(* IEC 61131-3 sources: plcassist-cli/packages/volt-lsp-iec/test-corpus/lenze-mid/Device/Plc Logic/Application/A70_MachineModuleSources/MM_MachineControl/02_subMain, 11 files *)

(* ---- SidecorrectionCalculation.fun ---- *)
FUNCTION SidecorrectionCalculation
VAR_INPUT
	iAnalogInputValue						: INT;
	iSetpoint								: INT;
	iCorrectionScale						: REAL;
	iLightValue								: INT;
	iDarkValue								: INT;
	iNoWrapperOffsetPercentage01Perc		: INT; //test5

END_VAR
VAR_OUTPUT
	oIntPercentage							: INT;
	oRealPercentage							: REAL;
	oCorrectionValue						: REAL;
	oDeviationNoWrapper						: REAL;
END_VAR
VAR

	tRealMeasuredValue						: REAL;
	tRealPercentage							: REAL;
	tRealSetpoint							: REAL;
	tWhiteValue								: DINT;
	tBrownValue								: DINT;
	tWidthLight_Dark						: DINT;
	tRealWidthLight_Dark					: REAL;
	tMeasuredWithOffset						: REAL;
	tRealBrownValue							: REAL;
	tRealNoWrapperOffsetPercentage			: REAL;

END_VAR

//Read out values for light and dark
tWhiteValue:=MOVE(iLightValue);
tBrownValue:=MOVE(iDarkValue);

//Calculate difference between light and dark value (light will be higher than dark)
tRealWidthLight_Dark:=TO_REAL(tWhiteValue-tBrownValue);
tRealBrownValue:=TO_REAL(tBrownValue);

//Measured value compensated with offset
tRealMeasuredValue:=TO_REAL(iAnalogInputValue);
tMeasuredWithOffset:=tRealMeasuredValue-tRealBrownValue;

//Calculation of the percentage
//"Measured value"/ Bandwidth
IF tRealWidthLight_Dark=0 THEN
	tRealWidthLight_Dark:=10;

END_IF
oRealPercentage:=(tMeasuredWithOffset/tRealWidthLight_Dark)*100;
oIntPercentage:=TO_INT(oRealPercentage);

//Calculation of the fault
//(act - set) * "correction scale"
tRealSetpoint:=TO_REAL(iSetpoint);
oCorrectionValue:=(oRealPercentage-tRealSetpoint)*iCorrectionScale;

//No wrapper detection
tRealNoWrapperOffsetPercentage:=TO_REAL(iNoWrapperOffsetPercentage01Perc);
oDeviationNoWrapper:=TO_INT(tRealNoWrapperOffsetPercentage*(tRealWidthLight_Dark/1000));

END_FUNCTION

(* ---- SpeedCalculationTrayfiller.fun ---- *)
FUNCTION SpeedCalculationTrayfiller
VAR_INPUT
END_VAR
VAR
	tInt: INT;
	tBool: BOOL;
END_VAR

NETWORK 0 LD TITLE: "NETWORK 1: Write setpoint speed in DB"
  // The speed of the trayfiller has to be higher then the speed of the dryer. In this way there is always an empty space at the startpostition of the trayfiller.
  LET en1 := ;
  IF en1 THEN tInt := (Mach1_Data.Drives.FeedForwardADS.Control.AutoSpeed + 30); END_IF
  LET en2 := en1;
  IF en2 THEN Mach1_Data.Drives.FeedForwardATF.Control.AutoSpeed := MOVE(tInt); END_IF
END_NETWORK
NETWORK 1 LD TITLE: "NETWORK 2: Activation + Runtime guard feed forward dryer/trayfiller"
  // Runtime calculation:
  // 1 cycle = 60s/rpm
  // speed = in 0.1 rpm -> 60s = 600 1/10s
  //
  // -> 1 cycle = 600/speed01
  // DINT cannot calculate this 600/1000 = 0.1 -> DINT=0
  // First multiply by 1000 (s -> ms)
  // 1cycle = (600*1000)/speed1
  // To give a little margin: add 500ms
  LET en1 := (Mach1.Genflags.DelayAfterSTO AND Mach1_Data.Drives.FeedForwardATF.Control.StartAuto AND NOT LST_InputsOutputs.I133_3_PROX_zero_position_transport_ATF);
  IF en1 THEN (Mach1_Data.Drives.FeedForwardATF.Control.AutoSpeed >= 10); END_IF
  Mach1.GenFlags.StopDriveDirect S= RuntimeGuard_V5_1_100(Mach1_Alarms, (Mach1_AuxData.TrayfillerActive AND Mach1_MIDS.IDB_TrayFiller.oFeedForwardMotor AND Mach1.Genflags.DelayAfterSTO AND (Mach1_AuxData.AllDrivesHomed OR NOT Mach1_AuxData.TrayfillerActive)), LST_General.AlwaysOff, en1, T#10S, Mach1.GenFlags.StartFlag, Mach1_Alarms.Alm051, Mach1.GenFlags.MinorAlarm, Mach1_AuxData.IEC_TIMERS.RuntimeGuardFeedforwardTrayfiller, oForwardGuarded => Mach1_Data.Drives.FeedForwardATF.Control.StartAuto);
END_NETWORK

END_FUNCTION

(* ---- Servo_LimitJog.fb ---- *)
FUNCTION_BLOCK Servo_LimitJog
VAR_INPUT
	iServoStatus 	: sUDT_ServoComm_Drive_Status;
	iServoControl 		: sUDT_ServoComm_Drive_Control;
END_VAR
VAR_OUTPUT
	oServoControl 		: sUDT_ServoComm_Drive_Control;
END_VAR
VAR
END_VAR
VAR_IN_OUT
	ioUDT_ServoDrive			: UDT_ServoDrive;
	ioUDT_JogLimitFree			: UDT_ServoJogLimitFree;
END_VAR

NETWORK 0 LD TITLE: "NETWORK 3 (p1): Check for limit switch"
  ioUDT_JogLimitFree.Status.Limit_Left_OK := iServoStatus.Spare1;
END_NETWORK
NETWORK 1 LD TITLE: "NETWORK 3 (p2): Check for limit switch"
  ioUDT_JogLimitFree.Status.Limit_Right_OK := iServoStatus.Spare2;
END_NETWORK
NETWORK 2 LD TITLE: "COPY previous control word to current controlword"
  LET en1 := ;
  IF en1 THEN
  EXECUTE
oServoControl:=iServoControl;
  END_EXECUTE
  END_IF
END_NETWORK
NETWORK 3 LD TITLE: "NETWORK 4 (p1): ControlToFreeLimitSwitches"
  oServoControl.Spare1 := (ioUDT_JogLimitFree.Status.Limit_Left_OK AND ioUDT_JogLimitFree.Control.Jog_LimitToLeft);
END_NETWORK
NETWORK 4 LD TITLE: "NETWORK 4 (p2): ControlToFreeLimitSwitches"
  oServoControl.Spare2 := (ioUDT_JogLimitFree.Status.Limit_Right_OK AND ioUDT_JogLimitFree.Control.Jog_LimitToRight);
END_NETWORK

END_FUNCTION_BLOCK

(* ---- WSM.fb ---- *)
FUNCTION_BLOCK WSM
VAR_INPUT
	EN: BOOL;
	iGenflags : UDT_GeneralFlags;
	iInit: BOOL;
	iTest_Prod: BOOL;
	iCleaning: BOOL;
	iBunchPresent: BOOL;
	iWrapperPresentForLeafCarrier: BOOL;
	iPhotocellWrapper: BOOL;
	iWaterLevelSensor: BOOL;
	iTakeOverCycle: BOOL;
	iTimeOutSupplyWrapper: TIME;
	iSprayTime: TIME;
	iDelayContSpraying: TIME;
	iScreenForOperatorSettingsActivated: BOOL;
	iManualSprayCycleReset: BOOL;
	iManualSprayCycleStart: BOOL;
	iManualSprayCycleStop: BOOL;
	iMaxNumberOfSprayPulses: INT;

END_VAR
VAR_OUTPUT
	ENO: BOOL;
	oVentilationMotor: BOOL;
	oPositionMotor: BOOL;
	oWindingMotor: BOOL;
	oSprayingValve: BOOL;
	oWaterLevelValve: BOOL;
	oFaultWaitingForWrapper: BOOL;
	oFaultNoWrapper: BOOL;
	oFaultPhotocellWrapper : BOOL;
END_VAR
VAR
	stOSN_TakeOverCycle: F_TRIG;
	TMR_TimeOutSupply: TON;
	TMR_TimeOutPhotocell: TON;
	stRePositionMotor: R_TRIG;
	stSprayCycleActive: BOOL;
	TMR_DelayContinuousSpraying: TON;
	TMR_SprayTime: TON;
	stManualSprayCycleStarted: BOOL;

	TMR_ManualSprayCycleIdle: TON;

END_VAR

VAR_IN_OUT
	ioEnableSpraying: BOOL;
	ioManualSprayCycleActualCount: INT;
	ioManualStartSupply: BOOL;
END_VAR
VAR RETAIN PERSISTENT
	stRestposition: BOOL;
	stSupplyWrapper: BOOL;
	stWrapperPresent: BOOL;
	stNoWrapper: BOOL;
	stPhotocellWrapperFault: BOOL;
	stFeedForward: BOOL;
END_VAR

NETWORK 0 LD TITLE: "DONE Network 2: State: Initialise"
  LET g8 := (iInit OR NOT iTest_Prod OR iCleaning OR ioManualStartSupply);
  stRestposition S= g8;
  LET g1 := g8;
  stSupplyWrapper R= g1;
  stWrapperPresent R= g1;
  stNoWrapper R= g1;
  stPhotocellWrapperFault R= g1;
END_NETWORK
NETWORK 1 LD TITLE: "DONE Network 3: State: Restposition"
  LET g1 := (stOSN_TakeOverCycle(CLK := iTakeOverCycle) AND stWrapperPresent);
  stRestposition S= g1;
  stWrapperPresent R= g1;
END_NETWORK
NETWORK 2 LD TITLE: "DONE Network 4: State: Supply wrapper"
  LET g1 := ((stRestposition AND ((iTest_Prod AND NOT iCleaning AND iBunchPresent AND NOT iTakeOverCycle AND (iGenFlags.RunMan OR iGenFlags.RunAuto)) OR ioManualStartSupply)) OR (stNoWrapper AND iGenFlags.StartFlag) OR (stPhotocellWrapperFault AND iGenFlags.StartFlag));
  stSupplyWrapper S= g1;
  stRestposition R= g1;
  stNoWrapper R= g1;
  stPhotocellWrapperFault R= g1;
  ioManualStartSupply R= g1;
END_NETWORK
NETWORK 3 LD TITLE: "DONE Network 5: State: Wrapper Present"
  LET g15 := (iWrapperPresentForLeafCarrier AND stSupplyWrapper);
  stWrapperPresent S= g15;
  LET en1 := g15;
  IF en1 THEN HMI_Var.Mach1.PRDWrapCurrentCntr := (1 + HMI_Var.Mach1.PRDWrapCurrentCntr); END_IF
  LET en2 := g15;
  IF en2 THEN HMI_Var.Mach1.PRDWrapDayCounter := (1 + HMI_Var.Mach1.PRDWrapDayCounter); END_IF
  stSupplyWrapper R= g15;
END_NETWORK
NETWORK 4 LD TITLE: "DONE Network 6: State: No Wrapper"
  LET g1 := TMR_TimeOutSupply(IN := (stSupplyWrapper AND stFeedForward), PT := iTimeOutSupplyWrapper);
  stNoWrapper S= g1;
  stSupplyWrapper R= g1;
END_NETWORK
NETWORK 5 LD TITLE: "DONE Network 7: State: Photocell wrapper fault"
  LET g1 := TMR_TimeOutPhotocell(IN := (stSupplyWrapper AND stFeedForward AND iPhotocellWrapper), PT := T#10S);
  stPhotocellWrapperFault S= g1;
  stSupplyWrapper R= g1;
END_NETWORK
NETWORK 6 LD TITLE: "DONE Network 8: Faults"
  LET g21 := True;
  oFaultWaitingForWrapper := (g21 AND stSupplyWrapper AND iTakeOverCycle);
  oFaultNoWrapper := (g21 AND stNoWrapper);
  oFaultPhotocellWrapper := (g21 AND stPhotocellWrapperFault);
END_NETWORK
NETWORK 7 LD TITLE: "DONE Network 9: Ventilation motor"
  oVentilationMotor := (iGenFlags.EnableAuxDrive AND iTest_Prod AND NOT iCleaning);
END_NETWORK
NETWORK 8 LD TITLE: "DONE Network 10:"
  LET g23 := (iGenFlags.EnableAuxDrive AND stSupplyWrapper AND NOT iGenFlags.StopFlag);
  stFeedForward := g23;
  oPositionMotor := g23;
END_NETWORK
NETWORK 9 LD TITLE: "DONE Network 11: Winding motor"
  oWindingMotor := (iGenFlags.EnableAuxDrive AND NOT iGenFlags.StopFlag AND iTest_Prod AND NOT iCleaning);
END_NETWORK
NETWORK 10 LD TITLE: "DONE Network 12: Start spray cycle"
  LET g46 := stFeedForward;
  stSprayCycleActive S= stRePositionMotor(CLK := g46);
  stSprayCycleActive S= TMR_DelayContinuousSpraying(IN := g46, PT := iDelayContSpraying);
END_NETWORK
NETWORK 11 LD TITLE: "DONE Network 13: Timing spray cycle"
  stSprayCycleActive R= (TMR_SprayTime(IN := stSprayCycleActive, PT := iSprayTime) AND NOT TMR_DelayContinuousSpraying.Q);
END_NETWORK
NETWORK 12 LD TITLE: "DONE Network 14: Spraying valve"
  oSprayingValve := (ioEnableSpraying AND stSprayCycleActive);
END_NETWORK
NETWORK 13 LD TITLE: "DONE Network 15: Automatic trigger of water"
  ioEnableSpraying S= (FALSE AND iGenFlags.EnablePneumEStop AND iWrapperPresentForLeafCarrier AND iTest_Prod AND NOT iCleaning);
END_NETWORK
NETWORK 14 LD TITLE: "DONE Network 16: Water level control"
  oWaterLevelValve := (ioEnableSpraying AND iWaterLevelSensor);
END_NETWORK
NETWORK 15 LD TITLE: "DONE Network 17: Manual spray cycle"
  LET g45 := iScreenForOperatorSettingsActivated;
  LET en1 := (g45 AND iManualSprayCycleReset);
  IF en1 THEN ioManualSprayCycleActualCount := MOVE(0); END_IF
  LET en2 := (g45 AND iGenFlags.EnablePneumEStop AND (iManualSprayCycleStart OR stManualSprayCycleStarted) AND NOT iManualSprayCycleStop AND NOT iManualSprayCycleReset);
  IF en2 THEN stManualSprayCycleStarted := (ioManualSprayCycleActualCount < iMaxNumberOfSprayPulses); END_IF
  LET en3 := TMR_ManualSprayCycleIdle(IN := (g45 AND stManualSprayCycleStarted AND NOT stSprayCycleActive), PT := T#300MS);
  IF en3 THEN ioManualSprayCycleActualCount := (ioManualSprayCycleActualCount + 1); END_IF
  stSprayCycleActive S= en3;
END_NETWORK
NETWORK 16 LD TITLE: "DONE Network 18: SAVE RLO"
  ENO := EN;
END_NETWORK

END_FUNCTION_BLOCK

(* ---- AHWF.prg ---- *)
PROGRAM AHWF
VAR
	tFaultWaitingForWrapper : BOOL;
	tFaultNoWrapper: BOOL;
	tFaultPhotocellWrapper: BOOL;
	tStartFastWinding: BOOL;
	tSupplyWrapper: BOOL;
	tSprayingValve: BOOL;
	ttest: BOOL;
	R_TrigStartPos: R_TRIG;
END_VAR

VAR
	IDB_WSM: WSM;
END_VAR

NETWORK 0 LD TITLE: "Network 1: Detection of wrapper (set and reset)"
  LET g10 := True;
  Mach1_AuxData.MemWrapperPassedUnderTheSensor S= (g10 AND LST_InputsOutputs.I101_0_Wrapper_present);
  LET g1 := (g10 AND NOT LST_InputsOutputs.I101_0_Wrapper_present AND Mach1_AuxData.MemWrapperPassedUnderTheSensor);
  Mach1_AuxData.MemWrapperPresentForLeafCarrier S= g1;
  Mach1_AuxData.MemWrapperDetected_ResetLimitedSpeed S= g1;
  LET en1 := g10;
  IF en1 THEN Mach1_AuxData.CamControls.TakeOverCycleStopPulse_CP.Start := MOVE(Mach1_Data.CamControls.TakeOverCycle_C.Stop); END_IF
  LET g2 := fc_CamC_CP_UDT(en1, HMI_Var.Mach1.Position, Mach1.GenFlags.Rotflag, Mach1_AuxData.CamControls.TakeOverCycleStopPulse_CP);
  Mach1_AuxData.MemWrapperPresentForLeafCarrier R= g2;
  Mach1_AuxData.MemWrapperPassedUnderTheSensor R= g2;
END_NETWORK
NETWORK 1 LD
  LET g1 := R_TrigStartPos(CLK := HMI_Var.HMI_AHWF_StartPos);
  Mach1_AuxData.MemWrapperPresentForLeafCarrier R= g1;
  Mach1_AuxData.MemWrapperPassedUnderTheSensor R= g1;
END_NETWORK
NETWORK 2 LD TITLE: "Network 2: FB for DTA"
  LET i1 := fc_dinttotime(Mach1_Data.Timers.TimeOutSupplyWrapper,2);
  LET i2 := fc_dinttotime(Mach1_Data.Timers.SprayPulseWidth,2);
  LET i3 := fc_dinttotime(Mach1_Data.Timers.DelayContSpraying,2);
  LET en1 := ;
  IF en1 THEN IDB_WSM(iGenflags := Mach1.GenFlags, iInit := LST_General.FirstCycle, iTest_Prod := HMI_Var.Test_Prod, iCleaning := HMI_Var.Btn_Cleaning, iBunchPresent := Mach1_AuxData.ShiftRegister.SR_bunch_present_position_1_JL, iWrapperPresentForLeafCarrier := (Mach1_AuxData.MemWrapperPresentForLeafCarrier AND NOT HMI_Var.HMI_AHWF_fast_winding), iPhotocellWrapper := (LST_InputsOutputs.I101_0_Wrapper_present AND NOT HMI_Var.HMI_AHWF_fast_winding), iWaterLevelSensor := LST_InputsOutputs.I101_3_Water_level_control, iTakeOverCycle := fc_CamC_CC_UDT(True, HMI_Var.Mach1.Position, Mach1_Data.CamControls.TakeOverCycle_C), iTimeOutSupplyWrapper := i1, iSprayTime := i2, iDelayContSpraying := i3, iScreenForOperatorSettingsActivated := Mach1_AuxData.ScreenForOperatorSettingsActivated, iManualSprayCycleReset := HMI_Var.Mach1.SprayReset, iManualSprayCycleStart := HMI_Var.Mach1.SprayStart, iManualSprayCycleStop := HMI_Var.Mach1.SprayStop, iMaxNumberOfSprayPulses := Mach1_Data.Settings.Ints.MaxNumberOfSprayPulses, ioEnableSpraying := HMI_Var.Btn_Spraying, ioManualSprayCycleActualCount := Mach1_Data.Settings.Ints.ActualNumberOfSprayPulses, ioManualStartSupply := HMI_Var.HMI_AHWF_StartPos, oPositionMotor => tSupplyWrapper, oSprayingValve => tSprayingValve, oWaterLevelValve => LST_InputsOutputs.Q101_1_PNV_Waterlevel_control, oFaultWaitingForWrapper => tFaultWaitingForWrapper, oFaultNoWrapper => tFaultNoWrapper, oFaultPhotocellWrapper => tFaultPhotocellWrapper); END_IF
  PneumValveTerminalSMC.Pos1B := (en1 AND Mach1.GenFlags.EnablePneumPressurised AND Mach1_Safety.Status.AllDoorsActuallyClosed AND tSprayingValve AND NOT Mach1_Alarms.Alm011);
END_NETWORK
NETWORK 3 LD TITLE: "Network 3: Wrapper faults"
  Mach1.GenFlags.StopDriveDirect S= (Alarms_V5_1_100(Mach1_Alarms, (Mach1.GenFlags.DelayAfterEmergStop AND HMI_Var.Test_Prod AND NOT HMI_Var.Btn_Cleaning AND tFaultWaitingForWrapper AND Mach1_AuxData.AllDrivesHomed), True, Mach1_Alarms.Alm076, Mach1.GenFlags.Warning) OR Alarms_V5_1_100(Mach1_Alarms, (Mach1.GenFlags.DelayAfterEmergStop AND HMI_Var.Test_Prod AND NOT HMI_Var.Btn_Cleaning AND tFaultNoWrapper AND Mach1_AuxData.AllDrivesHomed), Mach1.GenFlags.StartFlag, Mach1_Alarms.Alm043, Mach1.GenFlags.MinorAlarm) OR Alarms_V5_1_100(Mach1_Alarms, (Mach1.GenFlags.DelayAfterEmergStop AND HMI_Var.Test_Prod AND NOT HMI_Var.Btn_Cleaning AND NOT Mach1_Alarms.Alm045 AND tFaultPhotocellWrapper AND Mach1_AuxData.AllDrivesHomed), Mach1.GenFlags.StartFlag, Mach1_Alarms.Alm045, Mach1.GenFlags.MinorAlarm));
END_NETWORK
NETWORK 4 LD
END_NETWORK
NETWORK 5 LD TITLE: "TODO Network 4:"
  LET g328 := True;
  LET g329 := (g328 AND True);
  LET en1 := (g329 AND TRUE);
  IF en1 THEN Data_Exchange_Motion.FeedForwardWrapper.Control.VelUnit := MOVE(175); END_IF
  LET en2 := en1;
  IF en2 THEN Data_Exchange_Motion.FeedForwardWrapper.Control.DecUnit := MOVE(2000); END_IF
  LET en3 := en2;
  IF en3 THEN Data_Exchange_Motion.FeedForwardWrapper.Control.AccUnit := MOVE(750); END_IF
  LET en4 := en3;
  IF en4 THEN Data_Exchange_Motion.FeedForwardWrapper.Control.TorqueLimit := MOVE(100); END_IF
  LET g330 := (g329 AND HMI_Var.HMI_AHWF_fast_winding);
  tStartFastWinding := Mach1_AuxData.IEC_TIMERS.TON_StartFastWinding(IN := g330, PT := T#200MS);
  LET en5 := g330;
  IF en5 THEN Data_Exchange_Motion.FeedForwardWrapper.Control.VelUnit := MOVE(500); END_IF
  LET i1 := DINT_TO_LREAL(Mach1_Data.Settings.Dints.WrapperStopPosition)/10;
  LET en6 := g328;
  IF en6 THEN Data_Exchange_Motion.FeedForwardWrapper.Control.PosUnit := MOVE(i1); END_IF
  Data_Exchange_Motion.FeedForwardWrapper.Control.StartTouchprobePos := (g328 AND NOT HMI_Var.HMI_AHWF_positioningType AND NOT Mach1_Alarms.Alm056 AND mach1.Genflags.EnableAuxDrive AND (tSupplyWrapper OR tStartFastWinding OR (Data_Exchange_Motion.FeedForwardWrapper.Control.StartTouchprobePos AND NOT Data_Exchange_Motion.FeedForwardWrapper.Status.InPosition)));
  HMI_Var.HMI_AHWF_fast_winding R= Mach1_AuxData.Edge.OSP_StopFlag(CLK := (g328 AND (NOT Mach1_MIDS.FB_Mach1.iStop1 OR NOT Mach1_MIDS.FB_Mach1.iStop2 OR NOT Mach1_MIDS.FB_Mach1.iStop3 OR NOT Mach1_Safety.Status.AllDoorsActuallyClosed OR LST_InputsOutputs.I101_0_Wrapper_present)));
END_NETWORK
NETWORK 6 LD TITLE: "Network 5: Side correction"
  LET en1 := ;
  IF en1 THEN ??? := SideCorrection(); END_IF
END_NETWORK
NETWORK 7 LD TITLE: "Network 6: DTA-alarm: side limit reached"
  Mach1.GenFlags.StopDriveDirect S= (Alarms_V5_1_100(Mach1_Alarms, (Mach1_AuxData.Edge.OSP_LimitDTA_Reached(CLK := (Mach1_AuxData.MIDS_Active AND Mach1.GenFlags.DelayAfterEmergStop AND (NOT Mach1_Data.Drives.SideCorrection_FreeLimit.Status.Limit_Left_OK OR NOT Mach1_Data.Drives.SideCorrection_FreeLimit.Status.Limit_Right_OK))) AND Mach1_AuxData.AllDrivesHomed), Mach1.GenFlags.StartFlag, Mach1_Alarms.Alm057, Mach1.GenFlags.MinorAlarm) OR (LST_General.AlwaysOff AND Alarms_V5_1_100(Mach1_Alarms, (Mach1_AuxData.MIDS_Active AND Mach1.GenFlags.DelayAfterEmergStop AND (NOT Mach1_Data.Drives.SideCorrection_FreeLimit.Status.Limit_Left_OK OR NOT Mach1_Data.Drives.SideCorrection_FreeLimit.Status.Limit_Right_OK) AND Mach1_AuxData.AllDrivesHomed), Mach1.GenFlags.StartFlag, Mach1_Alarms.Alm074, Mach1.GenFlags.Warning)));
END_NETWORK
NETWORK 8 LD TITLE: "Network 7: Alarm: Water receptacle full"
  Mach1.GenFlags.StopDriveDirect S= Alarms_V5_1_100(Mach1_Alarms, (Mach1_AuxData.IEC_TIMERS.WaterReceptacleFull(IN := (Mach1_AuxData.MIDS_Active AND LST_InputsOutputs.I101_3_Water_level_control AND NOT Mach1_Alarms.Alm055), PT := T#5M) AND HMI_Var.Test_Prod AND HMI_Var.Btn_Spraying AND Mach1_AuxData.AllDrivesHomed), Mach1.GenFlags.StartFlag, Mach1_Alarms.Alm055, Mach1.GenFlags.MinorAlarm);
END_NETWORK

END_PROGRAM

(* ---- fc_CheckRegister.prg ---- *)
PROGRAM fc_CheckRegister
VAR
END_VAR

NETWORK 0 LD TITLE: "NETWORK 1: Shift CheckRegister"
  fc_ShiftRegister(db_CheckRegister.Positie);
END_NETWORK
NETWORK 1 LD TITLE: "NETWORK 2: Check for error in dryer"
  fc_CheckNumberOfErrorsRegister(db_CheckRegister.Positie, CTE.posCigarPresentOutfeed, Mach1_Data.Counters.MaxRepetitionNoCigarsDryer.SetValue, oError => db_CheckRegister.CheckRegisterError);
END_NETWORK

END_PROGRAM

(* ---- fc_Visualisation_HMI.prg ---- *)
PROGRAM fc_Visualisation_HMI
VAR_INPUT
END_VAR
VAR
	tbool: BOOL;
END_VAR

NETWORK 0 LD TITLE: "NETWORK 5: (P1) Visualisation - emergency stop"
  Alarms_V5_1_100(Mach1_Alarms, (Mach1_AuxData.MIDS_Active AND NOT Mach1_Safety.Status.Emergency_button01), True, Mach1_Alarms.Alm080, Mach1.GenFlags.warning);
END_NETWORK
NETWORK 1 LD TITLE: "NETWORK 5: (P2) Visualisation - emergency stop"
  Alarms_V5_1_100(Mach1_Alarms, (Mach1_AuxData.MIDS_Active AND NOT Mach1_Safety.Status.Emergency_button02), True, Mach1_Alarms.Alm081, Mach1.GenFlags.warning);
END_NETWORK
NETWORK 2 LD TITLE: "NETWORK 5: (P3) Visualisation - emergency stop"
  Alarms_V5_1_100(Mach1_Alarms, (Mach1_AuxData.MIDS_Active AND NOT Mach1_Safety.Status.Emergency_button04), True, Mach1_Alarms.Alm082, Mach1.GenFlags.warning);
END_NETWORK
NETWORK 3 LD TITLE: "DONE NETWORK 5 (p2): Visualisation - doors"
  tbool := (Alarms_V5_1_100(Mach1_Alarms, (Mach1_AuxData.MIDS_Active AND Mach1.Genflags.DelayAfterEmergStop AND NOT Mach1_Safety.Status.Door_switch01), True, Mach1_Alarms.Alm083, Mach1.GenFlags.warning) OR Alarms_V5_1_100(Mach1_Alarms, (Mach1_AuxData.MIDS_Active AND Mach1.Genflags.DelayAfterEmergStop AND NOT Mach1_Safety.Status.Door_switch02), True, Mach1_Alarms.Alm084, Mach1.GenFlags.warning) OR Alarms_V5_1_100(Mach1_Alarms, (Mach1_AuxData.MIDS_Active AND Mach1.Genflags.DelayAfterEmergStop AND NOT Mach1_Safety.Status.Door_switch03), True, Mach1_Alarms.Alm085, Mach1.GenFlags.warning) OR Alarms_V5_1_100(Mach1_Alarms, (Mach1_AuxData.MIDS_Active AND Mach1.Genflags.DelayAfterEmergStop AND NOT Mach1_Safety.Status.Door_switch04), True, Mach1_Alarms.Alm086, Mach1.GenFlags.warning) OR Alarms_V5_1_100(Mach1_Alarms, (Mach1_AuxData.MIDS_Active AND Mach1.Genflags.DelayAfterEmergStop AND NOT Mach1_Safety.Status.Door_switch05), True, Mach1_Alarms.Alm087, Mach1.GenFlags.warning));
END_NETWORK
NETWORK 4 LD
  tbool := (Alarms_V5_1_100(Mach1_Alarms, (Mach1_AuxData.MIDS_Active AND Mach1.Genflags.DelayAfterEmergStop AND NOT Mach1_Safety.Status.Door_switch06), True, Mach1_Alarms.Alm088, Mach1.GenFlags.warning) OR Alarms_V5_1_100(Mach1_Alarms, (Mach1_AuxData.MIDS_Active AND Mach1.Genflags.DelayAfterEmergStop AND NOT Mach1_Safety.Status.Door_switch07), True, Mach1_Alarms.Alm089, Mach1.GenFlags.warning) OR Alarms_V5_1_100(Mach1_Alarms, (Mach1_AuxData.MIDS_Active AND Mach1.Genflags.DelayAfterEmergStop AND NOT Mach1_Safety.Status.Door_switch08), True, Mach1_Alarms.Alm090, Mach1.GenFlags.warning) OR Alarms_V5_1_100(Mach1_Alarms, (Mach1_AuxData.MIDS_Active AND Mach1.Genflags.DelayAfterEmergStop AND NOT Mach1_Safety.Status.Door_switch09), True, Mach1_Alarms.Alm091, Mach1.GenFlags.warning) OR Alarms_V5_1_100(Mach1_Alarms, (Mach1_AuxData.MIDS_Active AND Mach1.Genflags.DelayAfterEmergStop AND NOT Mach1_Safety.Status.Door_switch10), True, Mach1_Alarms.Alm092, Mach1.GenFlags.warning));
END_NETWORK
NETWORK 5 LD
  tbool := (Alarms_V5_1_100(Mach1_Alarms, (Mach1_AuxData.MIDS_Active AND Mach1.Genflags.DelayAfterEmergStop AND NOT Mach1_Safety.Status.Door_switch14), True, Mach1_Alarms.Alm093, Mach1.GenFlags.warning) OR Alarms_V5_1_100(Mach1_Alarms, (Mach1_AuxData.MIDS_Active AND Mach1.Genflags.DelayAfterEmergStop AND NOT Mach1_Safety.Status.Door_switch15), True, Mach1_Alarms.Alm094, Mach1.GenFlags.warning) OR Alarms_V5_1_100(Mach1_Alarms, (Mach1_AuxData.MIDS_Active AND Mach1.Genflags.DelayAfterEmergStop AND NOT Mach1_Safety.Status.Door_switch16), True, Mach1_Alarms.Alm095, Mach1.GenFlags.warning) OR Alarms_V5_1_100(Mach1_Alarms, (Mach1_AuxData.MIDS_Active AND Mach1.Genflags.DelayAfterEmergStop AND NOT Mach1_Safety.Status.Door_switch11), True, Mach1_Alarms.Alm070, Mach1.GenFlags.warning) OR Alarms_V5_1_100(Mach1_Alarms, (Mach1_AuxData.MIDS_Active AND Mach1.Genflags.DelayAfterEmergStop AND NOT Mach1_Safety.Status.Door_switch12), True, Mach1_Alarms.Alm071, Mach1.GenFlags.warning));
END_NETWORK
NETWORK 6 LD
  Alarms_V5_1_100(Mach1_Alarms, (Mach1_AuxData.MIDS_Active AND Mach1.Genflags.DelayAfterEmergStop AND NOT Mach1_Safety.Status.Door_switch13), True, Mach1_Alarms.Alm072, Mach1.GenFlags.warning);
END_NETWORK
NETWORK 7 LD
  tbool := (Alarms_V5_1_100(Mach1_Alarms, (Mach1_AuxData.MIDS_Active AND Mach1.Genflags.DelayAfterEmergStop AND LST_InputsOutputs.I100_3_Selector_switch_auto_manual_OP0a), True, Mach1_Alarms.Alm018, Mach1.GenFlags.warning) OR Alarms_V5_1_100(Mach1_Alarms, (Mach1_AuxData.MIDS_Active AND Mach1.Genflags.DelayAfterEmergStop AND LST_InputsOutputs.I132_3_SW_Auto_Man), True, Mach1_Alarms.Alm019, Mach1.GenFlags.warning));
END_NETWORK
NETWORK 8 LD TITLE: "Reset of alarmlogging"
  LET en1 := HMI_Var.ResetAlarmLogging;
  IF en1 THEN HMI_Var.ResetAlarmLogging R= Alarms_ResetAlarmLogging(Mach1_Alarms); END_IF
END_NETWORK
NETWORK 9 LD TITLE: "Adding product counters"
  LET en1 := HMI_Var.Mach1.PRDCounterIncr;
  IF en1 THEN HMI_Var.Mach1.PRDTotalCounter := (HMI_Var.Mach1.PRDTotalCounter + 1); END_IF
  LET en2 := en1;
  IF en2 THEN HMI_Var.Mach1.PRDCigDayCounter := (HMI_Var.Mach1.PRDCigDayCounter + 1); END_IF
  LET en3 := en2;
  IF en3 THEN HMI_Var.Mach1.PRDCigCurrentCntr := (HMI_Var.Mach1.PRDCigCurrentCntr + 1); END_IF
  HMI_Var.Mach1.PRDCounterIncr R= en3;
END_NETWORK
NETWORK 10 LD TITLE: "Reset Day Counter"
  LET en1 := HMI_Var.Mach1.PRDDayCounterReset_01;
  IF en1 THEN HMI_Var.Mach1.PRDWrapDayCounter := MOVE(0); END_IF
  LET en2 := en1;
  IF en2 THEN HMI_Var.Mach1.PRDCigDayCounter := MOVE(0); END_IF
  HMI_Var.Mach1.PRDDayCounterReset_01 R= en2;
END_NETWORK
NETWORK 11 LD TITLE: "Reset Current Counter"
  LET en1 := HMI_Var.Mach1.PRDDayCounterReset;
  IF en1 THEN HMI_Var.Mach1.PRDWrapCurrentCntr := MOVE(0); END_IF
  LET en2 := en1;
  IF en2 THEN HMI_Var.Mach1.PRDCigCurrentCntr := MOVE(0); END_IF
  HMI_Var.Mach1.PRDDayCounterReset R= en2;
END_NETWORK
NETWORK 12 LD
  LET en1 := TRUE;
  IF en1 THEN PRG_AlarmsToDWord(); END_IF
END_NETWORK

END_PROGRAM

(* ---- MainDrive.prg ---- *)
PROGRAM MainDrive
VAR_INPUT
END_VAR
VAR
	tInt: INT;
	tMainDriveRun: BOOL;
	tMainDriveJog: BOOL;
END_VAR

VAR_OUTPUT
	oMainDriveRun: BOOL;
	oMainDriveJog: BOOL;
END_VAR

NETWORK 0 LD TITLE: "DONE NETWORK 1: Delay after doors closed"
  Mach1_AuxData.DelayAfterDoorsActuallyClosed := Mach1_AuxData.IEC_TIMERS.TON_DelayAfterDoorsClosed(IN := (Mach1.GenFlags.DelayAfterEmergStop AND Mach1_Safety.Status.AllDoorsActuallyClosed AND Mach1_Safety.Status.DoorsOK), PT := T#150MS);
END_NETWORK
NETWORK 1 LD TITLE: "DONE NETWORK 2: Activating main drive"
  LET g174 := TRUE;
  LET en1 := g174;
  IF en1 THEN tInt := MOVE(0); END_IF
  Mach1_AuxData.MemLowerSpeedBecauseOfNoWrapper R= (g174 AND NOT HMI_Var.Test_Prod);
  LET g175 := (g174 AND Mach1.GenFlags.EnableMainDrive AND Mach1.GenFlags.ConditionsReadyForOperation AND NOT Mach1.GenFlags.StopDriveDirect AND Mach1_AuxData.AllDrivesInLock);
  LET g176 := (g175 AND Mach1.GenFlags.RunAuto);
  LET g1 := g176;
  tMainDriveRun := g1;
  oMainDriveRun := g1;
  Mach1_Safety.Control.RequestAutoSpeed := g1;
  LET en2 := Mach1_AuxData.MemLowerSpeedBecauseOfNoWrapper;
  IF en2 THEN (Mach1_Data.AUTOSPEED <= 40); END_IF
  LET en3 := ((g176 AND (NOT Mach1_AuxData.MemLowerSpeedBecauseOfNoWrapper OR en2)) AND NOT HMI_Var.Btn_Cleaning);
  IF en3 THEN tInt := MOVE(Mach1_Data.AUTOSPEED); END_IF
  LET en4 := (g176 AND Mach1_AuxData.MemLowerSpeedBecauseOfNoWrapper);
  IF en4 THEN (Mach1_Data.AUTOSPEED > 40); END_IF
  LET en5 := (en4 AND NOT HMI_Var.Btn_Cleaning);
  IF en5 THEN tInt := MOVE(30); END_IF
  LET en6 := (g176 AND HMI_Var.Btn_Cleaning);
  IF en6 THEN tInt := MOVE(6); END_IF
  LET g177 := (g175 AND Mach1.GenFlags.RunMan);
  LET g2 := g177;
  tMainDriveJog := g2;
  oMainDriveJog := g2;
  Mach1_Safety.Control.RequestManSpeed := g2;
  LET en7 := g177;
  IF en7 THEN tInt := MOVE(Mach1_Data.MANUALSPEED); END_IF
  RPM_To_DriveSpeed(g174, tInt, oDriveSpeed => Mach1_Data.Drives.MainDrive_VM.Control.DriveMasterSpeed);
END_NETWORK
NETWORK 2 LD TITLE: "DONE NETWORK 3 : DriveIsRunning flag"
  LET g96 := TRUE;
  Mach1.GenFlags.StopDriveDirect R= g96;
  Mach1.GenFlags.DriveIsRunning := (g96 AND (tMainDriveRun OR tMainDriveJog));
  Mach1.GenFlags.DriveAtSpeed := Mach1_AuxData.IEC_TIMERS.TOFF_MainDriveAtProductionSpeed(IN := Mach1_AuxData.IEC_TIMERS.TON_MainDriveAtProductionSpeed(IN := (g96 AND tMainDriveRun), PT := T#200MS), PT := T#60MS);
END_NETWORK
NETWORK 3 LD TITLE: "DONE NETWORK 4: Alarm: Main drive blocked"
  LET en1 := Mach1_AuxData.IEC_TIMERS.TON_MainDriveBlocked(IN := oMainDriveRun, PT := T#12S);
  IF en1 THEN (HMI_Var.Mach1.ActualSpeed < 5); END_IF
  Mach1.GenFlags.StopDriveDirect S= (Alarms_V5_1_100(Mach1_Alarms, en1, Mach1.GenFlags.StartFlag, Mach1_Alarms.Alm040, Mach1.GenFlags.MinorAlarm) AND Mach1_Alarms.Alm040);
END_NETWORK
NETWORK 4 LD TITLE: "DONE NETWORK 5: Manual brakerelease" DISABLED
  LET g180 := TRUE;
  LST_InputsOutputs.Q101_0_REL_release_brake := (g180 AND Mach1_Alarms.Alm001 AND HMI_Var.ReleaseBrake);
  HMI_Var.ReleaseBrake R= (g180 AND (NOT Mach1_Alarms.Alm001 OR (Mach1_Alarms.Alm001 AND NOT Mach1.GenFlags.StartFlag)));
END_NETWORK

END_PROGRAM

(* ---- PRG_AlarmsToDWord.prg ---- *)
PROGRAM PRG_AlarmsToDWord
VAR
END_VAR

dwErrorWord1.0:=Mach1_Alarms.Alm001;
dwErrorWord1.1:=Mach1_Alarms.Alm002;
dwErrorWord1.2:=Mach1_Alarms.Alm003;
dwErrorWord1.3:=Mach1_Alarms.Alm004;
dwErrorWord1.4:=Mach1_Alarms.Alm005;
dwErrorWord1.5:=Mach1_Alarms.Alm006;
dwErrorWord1.6:=Mach1_Alarms.Alm007;
dwErrorWord1.7:=Mach1_Alarms.Alm008;
dwErrorWord1.8:=Mach1_Alarms.Alm009;
dwErrorWord1.9:=Mach1_Alarms.Alm010;
dwErrorWord1.10:=Mach1_Alarms.Alm011;
dwErrorWord1.11:=Mach1_Alarms.Alm012;
dwErrorWord1.12:=Mach1_Alarms.Alm013;
dwErrorWord1.13:=Mach1_Alarms.Alm014;
dwErrorWord1.14:=Mach1_Alarms.Alm015;
dwErrorWord1.15:=Mach1_Alarms.Alm016;
dwErrorWord1.16:=Mach1_Alarms.Alm017;
dwErrorWord1.17:=Mach1_Alarms.Alm018;
dwErrorWord1.18:=Mach1_Alarms.Alm019;
dwErrorWord1.19:=Mach1_Alarms.Alm020;
dwErrorWord1.20:=Mach1_Alarms.Alm021;
dwErrorWord1.21:=Mach1_Alarms.Alm022;
dwErrorWord1.22:=Mach1_Alarms.Alm023;
dwErrorWord1.23:=Mach1_Alarms.Alm024;
dwErrorWord1.24:=Mach1_Alarms.Alm025;
dwErrorWord1.25:=Mach1_Alarms.Alm026;
dwErrorWord1.26:=Mach1_Alarms.Alm027;
dwErrorWord1.27:=Mach1_Alarms.Alm028;
dwErrorWord1.28:=Mach1_Alarms.Alm029;
dwErrorWord1.29:=Mach1_Alarms.Alm030;
dwErrorWord1.30:=Mach1_Alarms.Alm031;
dwErrorWord1.31:=Mach1_Alarms.Alm032;

dwErrorWord2.0:=Mach1_Alarms.Alm033;
dwErrorWord2.1:=Mach1_Alarms.Alm034;
dwErrorWord2.2:=Mach1_Alarms.Alm035;
dwErrorWord2.3:=Mach1_Alarms.Alm036;
dwErrorWord2.4:=Mach1_Alarms.Alm037;
dwErrorWord2.5:=Mach1_Alarms.Alm038;
dwErrorWord2.6:=Mach1_Alarms.Alm039;
dwErrorWord2.7:=Mach1_Alarms.Alm040;
dwErrorWord2.8:=Mach1_Alarms.Alm041;
dwErrorWord2.9:=Mach1_Alarms.Alm042;
dwErrorWord2.10:=Mach1_Alarms.Alm043;
dwErrorWord2.11:=Mach1_Alarms.Alm044;
dwErrorWord2.12:=Mach1_Alarms.Alm045;
dwErrorWord2.13:=Mach1_Alarms.Alm046;
dwErrorWord2.14:=Mach1_Alarms.Alm047;
dwErrorWord2.15:=Mach1_Alarms.Alm048;
dwErrorWord2.16:=Mach1_Alarms.Alm049;
dwErrorWord2.17:=Mach1_Alarms.Alm050;
dwErrorWord2.18:=Mach1_Alarms.Alm051;
dwErrorWord2.19:=Mach1_Alarms.Alm052;
dwErrorWord2.20:=Mach1_Alarms.Alm053;
dwErrorWord2.21:=Mach1_Alarms.Alm054;
dwErrorWord2.22:=Mach1_Alarms.Alm055;
dwErrorWord2.23:=Mach1_Alarms.Alm056;
dwErrorWord2.24:=Mach1_Alarms.Alm057;
dwErrorWord2.25:=Mach1_Alarms.Alm058;
dwErrorWord2.26:=Mach1_Alarms.Alm059;
dwErrorWord2.27:=Mach1_Alarms.Alm060;
dwErrorWord2.28:=Mach1_Alarms.Alm061;
dwErrorWord2.29:=Mach1_Alarms.Alm062;
dwErrorWord2.30:=Mach1_Alarms.Alm063;
dwErrorWord2.31:=Mach1_Alarms.Alm064;

dwErrorWord3.0:=Mach1_Alarms.Alm065;
dwErrorWord3.1:=Mach1_Alarms.Alm066;
dwErrorWord3.2:=Mach1_Alarms.Alm067;
dwErrorWord3.3:=Mach1_Alarms.Alm068;
dwErrorWord3.4:=Mach1_Alarms.Alm069;
dwErrorWord3.5:=Mach1_Alarms.Alm070;
dwErrorWord3.6:=Mach1_Alarms.Alm071;
dwErrorWord3.7:=Mach1_Alarms.Alm072;
dwErrorWord3.8:=Mach1_Alarms.Alm073;
dwErrorWord3.9:=Mach1_Alarms.Alm074;
dwErrorWord3.10:=Mach1_Alarms.Alm075;
dwErrorWord3.11:=Mach1_Alarms.Alm076;
dwErrorWord3.12:=Mach1_Alarms.Alm077;
dwErrorWord3.13:=Mach1_Alarms.Alm078;
dwErrorWord3.14:=Mach1_Alarms.Alm079;
dwErrorWord3.15:=Mach1_Alarms.Alm080;
dwErrorWord3.16:=Mach1_Alarms.Alm081;
dwErrorWord3.17:=Mach1_Alarms.Alm082;
dwErrorWord3.18:=Mach1_Alarms.Alm083;
dwErrorWord3.19:=Mach1_Alarms.Alm084;
dwErrorWord3.20:=Mach1_Alarms.Alm085;
dwErrorWord3.21:=Mach1_Alarms.Alm086;
dwErrorWord3.22:=Mach1_Alarms.Alm087;
dwErrorWord3.23:=Mach1_Alarms.Alm088;
dwErrorWord3.24:=Mach1_Alarms.Alm089;
dwErrorWord3.25:=Mach1_Alarms.Alm090;
dwErrorWord3.26:=Mach1_Alarms.Alm091;
dwErrorWord3.27:=Mach1_Alarms.Alm092;
dwErrorWord3.28:=Mach1_Alarms.Alm093;
dwErrorWord3.29:=Mach1_Alarms.Alm094;
dwErrorWord3.30:=Mach1_Alarms.Alm095;
dwErrorWord3.31:=Mach1_Alarms.Alm096;

dwErrorWord4.0:=Mach1_Alarms.Alm097;
dwErrorWord4.1:=Mach1_Alarms.Alm098;
dwErrorWord4.2:=Mach1_Alarms.Alm099;
dwErrorWord4.3:=Mach1_Alarms.Alm100;

END_PROGRAM

(* ---- SideCorrection.prg ---- *)
PROGRAM SideCorrection
VAR_INPUT
END_VAR
VAR
	tCorrectionScale			: DINT;
	tCorrectionScaleReal		: REAL;
	tReal						: REAL;
	tDint						: DINT;
	tInt						: INT;

	tbool: BOOL;
END_VAR

NETWORK 0 LD TITLE: "Network 1: Averaging of sensorsignal"
  LET i1 := TO_INT(LST_InputsOutputs.IW340_LeafCoverageSensor);
  LET en1 := ;
  IF en1 THEN fc_MeanValue(20, True, i1, db_MeanValuesSideCorrectionSensor.MeasurementValues, oMeanValue => DB_Kantcorrectie.MeasuredValue); END_IF
END_NETWORK
NETWORK 1 LD
  LET g62 := TRUE;
  LET en1 := (g62 AND DB_Kantcorrectie.CopyMeasuredToDark);
  IF en1 THEN DB_Kantcorrectie.DarkValue := MOVE(DB_Kantcorrectie.MeasuredValue); END_IF
  DB_Kantcorrectie.CopyMeasuredToDark R= en1;
  LET en2 := (g62 AND DB_Kantcorrectie.CopyMeasuredToLight);
  IF en2 THEN DB_Kantcorrectie.LightValue := MOVE(DB_Kantcorrectie.MeasuredValue); END_IF
  DB_Kantcorrectie.CopyMeasuredToLight R= en2;
END_NETWORK
NETWORK 2 LD TITLE: "Network 2: Read out inputvalue and calculate correctionvalue"
  LET en1 := TRUE;
  IF en1 THEN tCorrectionScale := MOVE(Mach1_Data.Settings.Ints.SideCorrectionScaleFactor); END_IF
  LET en2 := en1;
  IF en2 THEN SidecorrectionCalculation(DB_Kantcorrectie.MeasuredValue, DB_Kantcorrectie.Setpoint, -1, DB_Kantcorrectie.LightValue, DB_Kantcorrectie.DarkValue, DB_Kantcorrectie.NoWrapperPercentage, oIntPercentage => DB_Kantcorrectie.Percentage10, oCorrectionValue => DB_Kantcorrectie.MeasuredValueReal, oDeviationNoWrapper => tReal); END_IF
  LET i1 := REAL_TO_INT(tReal);
  LET en3 := en2;
  IF en3 THEN DB_Kantcorrectie.DeviationNoWrapper := MOVE(i1); END_IF
END_NETWORK
NETWORK 3 LD TITLE: "Network 3: Determine side-correction value"
  LET g85 := fc_CamC_CP_UDT(, HMI_Var.Mach1.Position, Mach1.GenFlags.Rotflag, Mach1_Data.CamControls.MeasurementForSidecorrection_CP);
  LET en1 := (g85 AND Mach1_Data.Drives.SideCorrection_FreeLimit.Status.Limit_Left_OK AND Mach1_Data.Drives.SideCorrection_FreeLimit.Status.Limit_right_OK);
  IF en1 THEN DB_Kantcorrectie.CopiedValueReal := MOVE(DB_Kantcorrectie.MeasuredValueReal); END_IF
  LET en2 := en1;
  IF en2 THEN DB_Kantcorrectie.CopiedValueInt := MOVE(DB_Kantcorrectie.Percentage10); END_IF
  LET g86 := (g85 AND Mach1_AuxData.MemWrapperDetected_ResetLimitedSpeed);
  Mach1_AuxData.MemLowerSpeedBecauseOfNoWrapper R= g86;
  Mach1_AuxData.MemWrapperDetected_ResetLimitedSpeed R= g86;
  LET en3 := g85;
  IF en3 THEN DB_Kantcorrectie.NoWrapperValue := (DB_Kantcorrectie.LightValue - DB_Kantcorrectie.DeviationNoWrapper); END_IF
  LET en4 := en3;
  IF en4 THEN (LST_InputsOutputs.IW340_LeafCoverageSensor > DB_Kantcorrectie.NoWrapperValue); END_IF
  Mach1_AuxData.MemLowerSpeedBecauseOfNoWrapper S= (en4 AND HMI_Var.Test_Prod);
END_NETWORK
NETWORK 4 LD TITLE: "DONE Network 4: In case a limit switch is reached: overwrite values"
  LET g48 := True;
  LET en1 := (g48 AND NOT Mach1_Data.Drives.SideCorrection_FreeLimit.Status.Limit_Left_OK AND Mach1_Data.Drives.SideCorrection_FreeLimit.Status.Limit_Right_OK);
  IF en1 THEN DB_Kantcorrectie.CopiedValueReal := MOVE(-100.0); END_IF
  LET en2 := (g48 AND NOT Mach1_Data.Drives.SideCorrection_FreeLimit.Status.Limit_Right_OK AND Mach1_Data.Drives.SideCorrection_FreeLimit.Status.Limit_Left_OK);
  IF en2 THEN DB_Kantcorrectie.CopiedValueReal := MOVE(100.0); END_IF
  LET en3 := en2;
  IF en3 THEN tCorrectionScale := MOVE(-1); END_IF
  LET en4 := (g48 AND ((NOT Mach1_Data.Drives.SideCorrection_FreeLimit.Status.Limit_Left_OK AND NOT Mach1_Data.Drives.SideCorrection_FreeLimit.Status.Limit_Right_OK) OR NOT HMI_Var.Test_Prod OR Mach1_AuxData.MemLowerSpeedBecauseOfNoWrapper));
  IF en4 THEN DB_Kantcorrectie.CopiedValueReal := MOVE(0.0); END_IF
  LET en5 := en4;
  IF en5 THEN tCorrectionScale := MOVE(1); END_IF
END_NETWORK
NETWORK 5 LD TITLE: "DONE Network 5: Write side-correction values to the servo drive"
  LET en1 := ;
  IF en1 THEN
  EXECUTE
tReal:=DB_Kantcorrectie.CopiedValueReal*DINT_TO_REAL(tCorrectionScale);
Mach1_Data.Drives.SideCorrection.CAM.Y_Scale_Recipe:=REAL_TO_INT(tReal/(-1000));
  END_EXECUTE
  END_IF
END_NETWORK
NETWORK 6 LD TITLE: "DONE Network 6 : Manual adjustment of the sidecorrection"
  LET g56 := True;
  Mach1_Data.Drives.SideCorrection_FreeLimit.Control.Jog_LimitToLeft := (g56 AND Mach1_Data.Drives.SideCorrection_FreeLimit.Status.Limit_Left_OK AND HMI_Var.Mach1.DTA_PositioningLeft);
  Mach1_Data.Drives.SideCorrection_FreeLimit.Control.Jog_LimitToRight := (g56 AND Mach1_Data.Drives.SideCorrection_FreeLimit.Status.Limit_Right_OK AND HMI_Var.Mach1.DTA_PositioningRight);
END_NETWORK

END_PROGRAM

(* ---- SpeedCalculationDryer.prg ---- *)
PROGRAM SpeedCalculationDryer
VAR_INPUT
END_VAR
VAR
	TempI: INT;
	cor_DenumI: INT:=1;
	cor_NumI: INT:=1;
	cor_DenumDI: DINT:=1;
	cor_NumDI: DINT:=1;
	Speed01rpm: INT;
	tSetHighSpeedCycles : BOOL;
	cor_Const: INT;
	R_TRIG_0: R_TRIG;
	MainDrive_AutoSpeed01rpm: INT;
	Mach_ActSpeed_Rpm01:INT;
	devAngle: INT;

END_VAR

NETWORK 0 LD TITLE: "NETWORK 1 : Speed control transport system dryer"
  LET g185 := True;
  LET en1 := g185;
  IF en1 THEN TempI := MOVE(0); END_IF
  LET en2 := g185;
  IF en2 THEN MainDrive_AutoSpeed01rpm := (Mach1_Data.AUTOSPEED * 10); END_IF
  LET en3 := g185;
  IF en3 THEN Droger_Data.Cor_denumerator := MOVE(MainDrive_AutoSpeed01rpm); END_IF
  LET g186 := (g185 AND True);
  LET en4 := (Mach1_AuxData.IEC_TIMERS.TON_DelayIdling(IN := (g186 AND NOT Mach1.GenFlags.DriveIsRunning), PT := T#500MS) AND NOT Mach1_Alarms.Alm049);
  IF en4 THEN Mach_ActSpeed_Rpm01 := MOVE(MainDrive_AutoSpeed01rpm); END_IF
  LET en5 := en4;
  IF en5 THEN Droger_Data.Cor_numerator := MOVE(MainDrive_AutoSpeed01rpm); END_IF
  LET en6 := (g186 AND (Mach1.GenFlags.DriveIsRunning OR NOT Mach1_AuxData.IEC_TIMERS.TON_DelayIdling.Q));
  IF en6 THEN Mach_ActSpeed_Rpm01 := MOVE(HMI_Var.Mach1.ActualSpeed*10); END_IF
  LET g187 := (g186 AND True);
  LET g188 := (g187 AND Trayfiller_Data.commInterface.HoldFeedFwd);
  LET en7 := (g188 AND (LST_InputsOutputs.I133_1_PROX_zero_position_transport_ADS OR Mach1_AuxData.ADS_StopOnZeroPulse));
  IF en7 THEN Droger_Data.Cor_numerator := MOVE(750); END_IF
  LET en8 := Mach1_AuxData.Edge.Osr_SetCounter(CLK := (g188 AND Trayfiller_Data.commInterface.Permission));
  IF en8 THEN Mach1_AuxData.CounterHighSpeedATF_ADS := MOVE(5); END_IF
  LET en9 := (g187 AND Trayfiller_Data.commInterface.Permission);
  IF en9 THEN (Mach1_AuxData.CounterHighSpeedATF_ADS <> 0); END_IF
  LET en10 := en9;
  IF en10 THEN Droger_Data.Cor_numerator := (Mach1_Data.AUTOSPEED * 13); END_IF
  LET en11 := g186;
  IF en11 THEN
  EXECUTE
cor_NumDI:=Droger_Data.Cor_numerator;
cor_DenumDI:=Droger_Data.Cor_denumerator;
//cor_NumDI:=1;
//cor_DenumDI:=1;
HMI_Var.Mach1.ActualSpeedDryer:=(Mach_ActSpeed_Rpm01*cor_numDI)/cor_denumdi;
Mach1_Data.Drives.FeedForwardADS.Control.AutoSpeed:=REAL_TO_INT(0.9*dint_to_real(HMI_Var.Mach1.ActualSpeedDryer)*6/10);
  END_EXECUTE
  END_IF
END_NETWORK
NETWORK 1 LD TITLE: "NETWORK 2: Deviation calculation of sync point, transport system trayfiller"
  // Principle: It's better to accelerate the drive then to decelerate, because otherwise cigars could be missed.
  // So that is why the deceleration should be kept short, by trial and error the optimum point is 60degrees (difference between setpoint and actual point).
  // dev: [0-60]: dec.
  // dev: ]60-360]: acc.
  //
  // Numerator = (Act_syncpos -/- Gew_syncpos) + Cte
  // Cte=little bit slower then the value for the set speed. (If the mid-s rotates 100rpm (value=1000), then this value should be a little less (e.g 99,8rpm).
  //         This way, the system lags a little bit, and therefor needs to accelerate (which is beter). If the system leads, then it needs to decel. (which is not ideal)
  //
  // Uit metingen is gebleken dat de optimale synchronisatiepositie op 60 graden
  // ligt.
  //
  // correctie  -60     0     60     120    180    240    300
  //             |------|------|------|------|------|------|--
  // encoder     0     60     120    180    240    300    360
  //
  // Om de ingestelde synchronisatiepositie te verschuiven naar het optimale window
  // van -60..300 wordt de correctiefactor gecorrigeerd:
  //  - indien correctie < -60 dan 360 erbij optellen
  //  - indien correctie > 300 dan 360 eraf tellen
  LET en1 := Mach1.GenFlags.DriveIsRunning;
  IF en1 THEN devAngle := (Droger_Data.Act_sync_pos - Droger_Data.set_sync_pos); END_IF
  LET en2 := en1;
  IF en2 THEN cor_Const := (MainDrive_AutoSpeed01rpm - 2); END_IF
  LET en3 := en2;
  IF en3 THEN Droger_Data.Cor_numerator := (devAngle + cor_Const); END_IF
  LET g4 := en3;
  LET en4 := g4;
  IF en4 THEN (devAngle < -60); END_IF
  LET en5 := en4;
  IF en5 THEN Droger_Data.Cor_numerator := (Droger_Data.Cor_numerator + 360); END_IF
  LET en6 := g4;
  IF en6 THEN (devAngle > 300); END_IF
  LET en7 := en6;
  IF en7 THEN Droger_Data.Cor_numerator := (Droger_Data.Cor_numerator - 360); END_IF
END_NETWORK
NETWORK 2 LD
  LET g0 := R_TRIG_0(CLK := LST_InputsOutputs.I133_1_PROX_zero_position_transport_ADS);
  LET en1 := g0;
  IF en1 THEN Droger_Data.Act_sync_pos := MOVE(HMI_Var.Mach1.Position); END_IF
  LET en2 := g0;
  IF en2 THEN Droger_Data.set_sync_pos := MOVE(Mach1_Data.CamControls.FeedforwardDryer_CP.Start); END_IF
  LET en3 := g0;
  IF en3 THEN (Mach1_AuxData.CounterHighSpeedATF_ADS > 0); END_IF
  LET en4 := en3;
  IF en4 THEN Mach1_AuxData.CounterHighSpeedATF_ADS := (Mach1_AuxData.CounterHighSpeedATF_ADS - 1); END_IF
END_NETWORK

END_PROGRAM
